// TIA Portal V20 export
DATA_BLOCK "OP1_DB"   // DB50
// stored: AutoNumber false, InstanceOfName OP1, InstanceOfType FB
"OP1"
   // VAR
   //    CONTROL_MAN : Struct
   //       kar_work : Bool;
   //       kar_home : Bool;
   //       zarazka_work : Bool;
   //       zarazka_home : Bool;
   //       B4 : Bool;
   //       B5 : Bool;
   //       B6 : Bool;
   //       B7 : Bool;
   //       B8 : Bool;
   //       B9 : Bool;
   //       odfuk_1 : Bool;
   //       odfuk_2 : Bool;
   //       B12 : Bool;
   //       B13 : Bool;
   //       B14 : Bool;
   //       B15 : Bool;
   //       B16 : Bool;
   //       B17 : Bool;
   //       B18 : Bool;
   //       B19 : Bool;
   //       B20 : Bool;
   //       B21 : Bool;
   //       B22 : Bool;
   //       B23 : Bool;
   //       B24 : Bool;
   //       B25 : Bool;
   //       B26 : Bool;
   //       B27 : Bool;
   //       B28 : Bool;
   //       B29 : Bool;
   //       B30 : Bool;
   //       B31 : Bool;
   //    END_STRUCT;
   //    CONTROL_AUTOMAT : Struct
   //       KAR_WORK : Bool;
   //       KAR_HOME : Bool;
   //       ZARAZKA_WORK : Bool;
   //       ZARAZKA_HOME : Bool;
   //       B4 : Bool;
   //       B5 : Bool;
   //       B6 : Bool;
   //       B7 : Bool;
   //       B8 : Bool;
   //       B9 : Bool;
   //       odfuk_1 : Bool;
   //       odfuk_2 : Bool;
   //       B12 : Bool;
   //       B13 : Bool;
   //       B14 : Bool;
   //       B15 : Bool;
   //       B16 : Bool;
   //       B17 : Bool;
   //       B18 : Bool;
   //       B19 : Bool;
   //       B20 : Bool;
   //       B21 : Bool;
   //       B22 : Bool;
   //       B23 : Bool;
   //       B24 : Bool;
   //       B25 : Bool;
   //       B26 : Bool;
   //       B27 : Bool;
   //       B28 : Bool;
   //       B29 : Bool;
   //       B30 : Bool;
   //       B31 : Bool;
   //    END_STRUCT;
   //    SENSORS : Struct
   //       prechod_1 : Bool;
   //       prechod_1_neg : Bool;
   //       kontrola : Bool;
   //       kontrola_neg : Bool;
   //       prechod_2 : Bool;
   //       Prechod_2_neg : Bool;
   //       Pozice_vyrazovace : Bool;
   //       Pozice_vyrazovace_neg : Bool;
   //       Pozice_pistu : Bool;
   //       Pozice_pistu_neg : Bool;
   //       s10 : Bool;
   //       s11 : Bool;
   //       s12 : Bool;
   //       s13 : Bool;
   //       s14 : Bool;
   //       s15 : Bool;
   //       s16 : Bool;
   //       s17 : Bool;
   //       s18 : Bool;
   //       s19 : Bool;
   //       s20 : Bool;
   //       s21 : Bool;
   //       s22 : Bool;
   //       s23 : Bool;
   //       s24 : Bool;
   //       s25 : Bool;
   //       s26 : Bool;
   //       s27 : Bool;
   //       s28 : Bool;
   //       s29 : Bool;
   //       s30 : Bool;
   //       s31 : Bool;
   //    END_STRUCT;
   //    SENSORS_1 : Struct
   //       S0 : Bool;
   //       S1 : Bool;
   //       S2 : Bool;
   //       S3 : Bool;
   //       S4 : Bool;
   //       S5 : Bool;
   //       S6 : Bool;
   //       S7 : Bool;
   //       S8 : Bool;
   //       S9 : Bool;
   //       SESTAVA_NENI_OTOCENA : Bool;
   //       SESTAVA_JE_OTOCENA : Bool;
   //       S12 : Bool;
   //       S13 : Bool;
   //       S14 : Bool;
   //       S15 : Bool;
   //       S16 : Bool;
   //       S17 : Bool;
   //       S18 : Bool;
   //       S19 : Bool;
   //       S20 : Bool;
   //       S21 : Bool;
   //       S22 : Bool;
   //       S23 : Bool;
   //       S24 : Bool;
   //       S25 : Bool;
   //       S26 : Bool;
   //       S27 : Bool;
   //       S28 : Bool;
   //       S29 : Bool;
   //       S30 : Bool;
   //       l_3_neg : Bool;
   //    END_STRUCT;
   //    S_0 : "SENSOR";
   //    S_1 : "SENSOR";
   //    S_2 { S7_SetPoint := 'True'} : "SENSOR";
   //    S_3 { S7_SetPoint := 'True'} : "SENSOR";
   //    S_4 { S7_SetPoint := 'True'} : "SENSOR";
   //    S_5 { S7_SetPoint := 'True'} : "SENSOR";
   //    S_6 { S7_SetPoint := 'True'} : "SENSOR";
   //    M_karusel : "MOTOR_CONTROL_BLOCK";
   //    M_zarazka { S7_SetPoint := 'True'} : "MOTOR_CONTROL_BLOCK";
   //    M_CLONA { S7_SetPoint := 'True'} : "MOTOR_CONTROL_BLOCK";
   //    SQCR { S7_SetPoint := 'True'} : Int;
   //    hmi_sqcr : Int;
   //    TRIG : Struct
   //       inicial_ok_op : Bool;
   //       DSSAD : Bool;
   //       INICIALIZACE_PROBEHLA : Bool;
   //       trig_dil : Bool;
   //       p_trig_control_tcon : Bool;
   //       T6 : Bool;
   //       SPUST_OP_4 : Bool;
   //       vlez_do_zavory_pri_rotaci : Bool;
   //       START_INICIAL_OP2 : Bool;
   //       START_INICIAL_OP3 : Bool;
   //       spust_odsavani : Bool;
   //       VYPRAZNI_OK_OP_2_A : Bool;
   //       VYPRAZNI_NOK_OP_2_A : Bool;
   //       VYPRAZDNI_OK_OP_3_B : Bool;
   //       VYPRAZDNI_NOK_OP_3_B : Bool;
   //       RESET_NCODER : Bool;
   //       op_1_ready : Bool;
   //    END_STRUCT;
   //    MEMOR : Struct
   //       n_trig_vypnuti : Bool;
   //       M1 : Bool;
   //       M2 : Bool;
   //       M3 : Bool;
   //       M4 : Bool;
   //       p_trig_odavacka : Bool;
   //       M6 : Bool;
   //       M7 : Bool;
   //       M8 : Bool;
   //       M9 : Bool;
   //       M10 : Bool;
   //       M11 : Bool;
   //       RESET_ERROR : Bool;
   //       vyrazeni_pamet : Bool;
   //       M14 : Bool;
   //       M15 : Bool;
   //       SETOVANI_START : Bool;
   //       M17 : Bool;
   //       p_trig_pamet_1 : Bool;
   //       p_trig_pamet_2 : Bool;
   //       p_trig_pamet_3 : Bool;
   //       p_trig_pamet_4 : Bool;
   //       p_trig_pamet_5 : Bool;
   //       p_trig_pamet_6 : Bool;
   //       p_trig_pamet_7 : Bool;
   //       p_trig_pamet_8 : Bool;
   //       p_trig_pamet_9 : Bool;
   //       p_trig_pamet_10 : Bool;
   //       p_trig_vyrad : Bool;
   //       p_Trig_cisteni_pozice : Bool;
   //       p_trig_citac : Bool;
   //       N_TRIG_SAFETY : Bool;
   //       P_TRIG_RESET_POZICE : Bool;
   //       M33 : Bool;
   //       start_caklu : Bool;
   //       M35 : Bool;
   //       M36 : Bool;
   //       M37 : Bool;
   //       M38 : Bool;
   //       M39 : Bool;
   //       ALARM_GLOBAL : Bool;
   //       M41 : Bool;
   //       M42 : Bool;
   //       M43 : Bool;
   //       M44 : Bool;
   //       M45 : Bool;
   //       M46 : Bool;
   //       M47 : Bool;
   //       M48 : Bool;
   //       M49 : Bool;
   //       wrong_p_trig : Bool;
   //       alarm_p_trig : Bool;
   //       M52 : Bool;
   //       M53 : Bool;
   //       M54 : Bool;
   //       M55 : Bool;
   //       M56 : Bool;
   //       M57 : Bool;
   //       M58 : Bool;
   //       M59 : Bool;
   //       M60 : Bool;
   //       M61 : Bool;
   //       M62 : Bool;
   //       M63 : Bool;
   //    END_STRUCT;
   //    "TIMER" : Struct
   //       TIMER_0 : IEC_TIMER;
   //       TIMER_VACUUM_CLEANER : IEC_TIMER;
   //       TIMER_DELAY_RESET_EXECUTE : IEC_TIMER;
   //       TIMER_3 : IEC_TIMER;
   //       TIMER_4 : IEC_TIMER;
   //       air : IEC_TIMER;
   //       TIMER_6 : IEC_TIMER;
   //       TIMER_7 : IEC_TIMER;
   //    END_STRUCT;
   //    HMI : Struct
   //       povoleni_volby_receptu : Bool;
   //       "svetlo_on/off" : Bool;
   //       ALARM_VIDITELNOST : Bool;
   //       hmi_3 : Bool;
   //       hmi_4 : Bool;
   //       reset_fronty : Bool;
   //       hmi_6 : Bool;
   //       hmi_7 : Bool;
   //       hmi_8 : Bool;
   //       hmi_9 : Bool;
   //       hmi_10 : Bool;
   //       hmi_11 : Bool;
   //       hmi_12 : Bool;
   //       hmi_13 : Bool;
   //       hmi_14 : Bool;
   //       hmi_15 : Bool;
   //    END_STRUCT;
   //    STRING_0 : String[1];
   //    array_chyb_ctec : Array[1..16] of Bool;
   //    zpracovani_dat { ExternalAccessible := 'False'; ExternalVisible := 'False'; ExternalWritable := 'False'} : Array[1..1] of Struct
   //       prenaseny_text : String[100];
   //       balik_den : Int;
   //       vyrazeni : Bool;
   //    END_STRUCT;
   //    aktual_kusy : Int;
   //    i : Int;
   //    q : Int;
   //    pocet_znaku_string_kamera : Int;
   //    ocekavany_text : String[100];
   //    format_etiketa_ok : Bool;
   //    Kamera : Struct
   //       s2_pamet : Bool;
   //       s2_nabeh : Bool;
   //       sber_aktivni : Bool;
   //       prijato_etiketa : Bool;
   //       prijato_folie_l : Bool;
   //       prijato_folie_p : Bool;
   //       ok_etiketa : Bool;
   //       ok_folie_l : Bool;
   //       ok_folie_p : Bool;
   //       vyradit : Bool;
   //       fronta_plna : Bool;
   //       bypass_ocr : Bool := false;
   //       last_id_etiketa : Word;
   //       last_id_folie_l : Word;
   //       last_id_folie_p : Word;
   //       balik_den : Int;
   //       idx : Int;
   //       pocet : Int;
   //       text_etiketa : String[100];
   //       timeout_sberu : Time;
   //       kontrola_tridirny : Bool;
   //       tridirna_ok : Bool;
   //    END_STRUCT;
   //    Vyrazeni : Struct
   //       s4_pamet : Bool;
   //       s4_nabeh : Bool;
   //       aktivni : Bool;
   //       vyradit : Bool;
   //       chyba_bez_dat : Bool;
   //       chyba_pist : Bool;
   //       max_puls : Time;
   //       vyrazovac_pripojen : Bool;
   //       alarm_nok_balik : Bool;
   //       posledni_nok_balik : Int;
   //       posledni_nok_text : String[100];
   //       pocet_nok : DInt;
   //       pocet_bez_dat : DInt;
   //       majak_tp : TP_TIME;
   //       majak { S7_SetPoint := 'True'} : Bool;
   //    END_STRUCT;
   //    Kam_Etiketa_Job : Struct
   //       krok : Int;
   //       pozadovany : Int;
   //       odesli_pamet : Bool;
   //       aktivni : Bool;
   //       chyba : Bool;
   //       chyba_kod : Word;
   //       nesouhlasi : Bool;
   //       timeout : Time;
   //    END_STRUCT;
   //    Test_tp_ka12 : TP_TIME;
   // END_VAR
BEGIN
END_DATA_BLOCK
